// Durée du cycle de la tâche courante en ms (docs/04 § 2)
FUNCTION F_CycleMs : LREAL
VAR
    nTask : DINT;
END_VAR

nTask := GETCURTASKINDEXEX();
F_CycleMs := UDINT_TO_LREAL(TwinCAT_SystemInfoVarList._TaskInfo[nTask].CycleTime) / 10000.0;

END_FUNCTION

(* stored: Version 1.1.0.1, ProductVersion 3.1.4024.12
   POU F_CycleMs: Id {d9114e1e-e081-56a8-b5e9-83cd581664aa}, SpecialFunc None *)
